(* Logix 5000 project; controller R400_500_XLS vendor 1 type 14 code 216 rev 31.11; software revision 31.01; part 11 of 32 *)
(* tags used below, declared in another part *)
   CalCond : SINT;
   CalFrinseCond : SINT;
   CalibCondCnt : SINT;
   CalibData : UDT_SCALE[8];
   CalibFrinseCondCnt : SINT;
   CalibIndex : DINT;   // Calibration Pointer
   CalibPressCnt : SINT;
   CalPressure : SINT;
   DX_div_100 : REAL;
   M : DINT[5];   // Memory Bits
   ONS_FC86 : DINT;
   rBuffer : REAL[4];
   Supervisor : DINT;
   ChemCond : REAL;
   FinalRinseCond : REAL;
   I_Chem_Cond : DINT;   // Chemical water conductivity
   I_Final_Rinse_Cond : DINT;   // Final rinse water conductivity
   I_Pump_Press : DINT;   // Recirculation pump pressure
   Msg_CalibChem : SINT;
   Msg_CalibFrinse : SINT;
   Msg_CalibPress : SINT;
   Msg_EditCalib : SINT;   // Screen 103 Msg Display
   NumInput : UDT_NUMERIC_INPUT[65];   // Numeric input
   NumInputReal : UDT_NUMERIC_INPUT_REAL[17];
   PmpPres : REAL;
   PressureUnit : BOOL;   // Pressure Unit 0=PSIG 1=BAR
   Screen_Ctrl : DINT;   // PLC Screen Request
   Tpb : DINT[11];
   TpbImage : DINT[11];
   Unit : Hrdwre;   // Unit Configuration
(* MainProgram, continued *)

ROUTINE SPV_10_ANALOG_CHANNEL_CALIBRATION   (* ladder *)
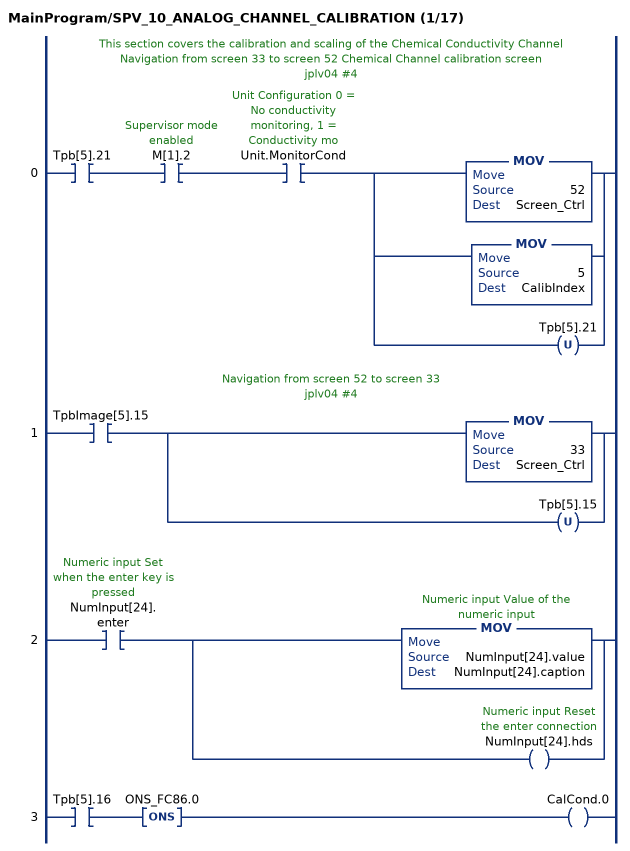
   // This section covers the calibration and scaling of the Chemical Conductivity Channel
   // Navigation from screen 33 to screen 52 Chemical Channel calibration screen
   // jplv04 #4
   0: XIC(Tpb[5].21)XIC(M[1].2)XIC(Unit.MonitorCond)[MOV(52,Screen_Ctrl) ,MOV(5,CalibIndex) ,OTU(Tpb[5].21) ];
   // Navigation from screen 52 to screen 33
   // jplv04 #4
   1: XIC(TpbImage[5].15)[MOV(33,Screen_Ctrl) ,OTU(Tpb[5].15) ];
   2: XIC(NumInput[24].enter)[MOV(NumInput[24].value,NumInput[24].caption) ,OTE(NumInput[24].hds) ];
   3: XIC(Tpb[5].16)ONS(ONS_FC86.0)OTE(CalCond.0);
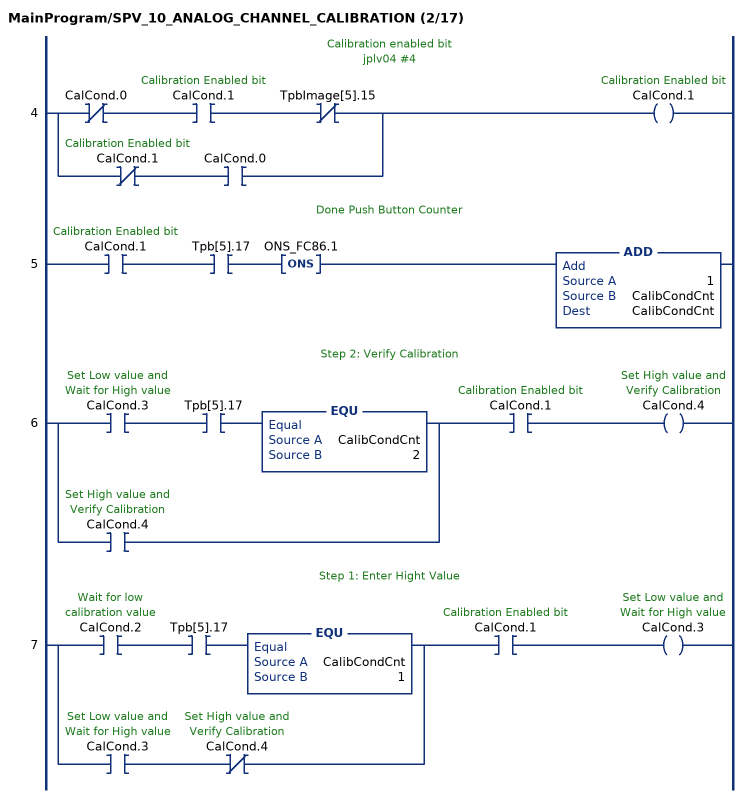
   // Calibration enabled bit
   // jplv04 #4
   4: [XIO(CalCond.0) XIC(CalCond.1) XIO(TpbImage[5].15) ,XIO(CalCond.1) XIC(CalCond.0) ]OTE(CalCond.1);
   // Done Push Button Counter
   5: XIC(CalCond.1)XIC(Tpb[5].17)ONS(ONS_FC86.1)ADD(1,CalibCondCnt,CalibCondCnt);
   // Step 2: Verify Calibration
   6: [XIC(CalCond.3) XIC(Tpb[5].17) EQU(CalibCondCnt,2) ,XIC(CalCond.4) ]XIC(CalCond.1)OTE(CalCond.4);
   // Step 1: Enter Hight Value
   7: [XIC(CalCond.2) XIC(Tpb[5].17) EQU(CalibCondCnt,1) ,XIC(CalCond.3) XIO(CalCond.4) ]XIC(CalCond.1)OTE(CalCond.3);
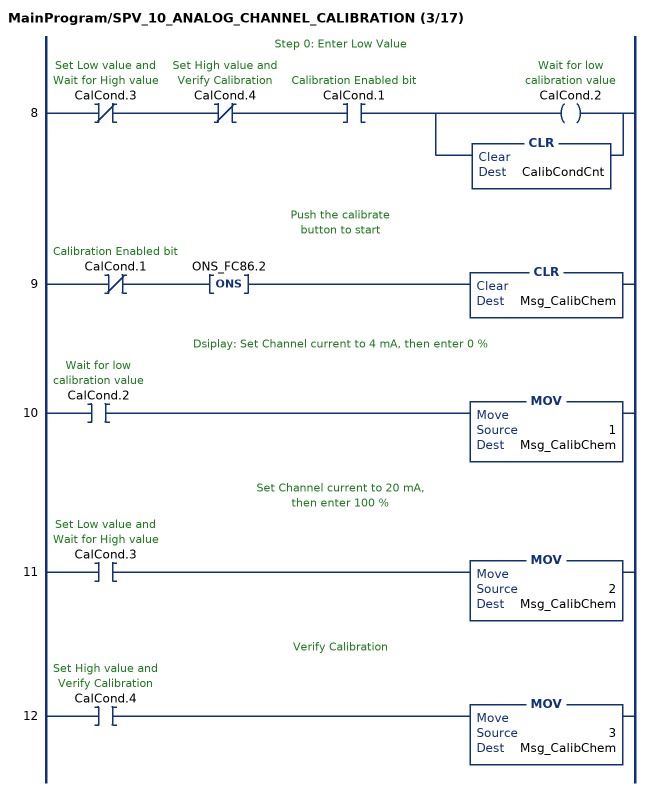
   // Step 0: Enter Low Value
   8: XIO(CalCond.3)XIO(CalCond.4)XIC(CalCond.1)[OTE(CalCond.2) ,CLR(CalibCondCnt) ];
   // Push the calibrate
   // button to start
   9: XIO(CalCond.1)ONS(ONS_FC86.2)CLR(Msg_CalibChem);
   // Dsiplay: Set Channel current to 4 mA, then enter 0 %
   10: XIC(CalCond.2)MOV(1,Msg_CalibChem);
   // Set Channel current to 20 mA,
   // then enter 100 %
   11: XIC(CalCond.3)MOV(2,Msg_CalibChem);
   // Verify Calibration
   12: XIC(CalCond.4)MOV(3,Msg_CalibChem);
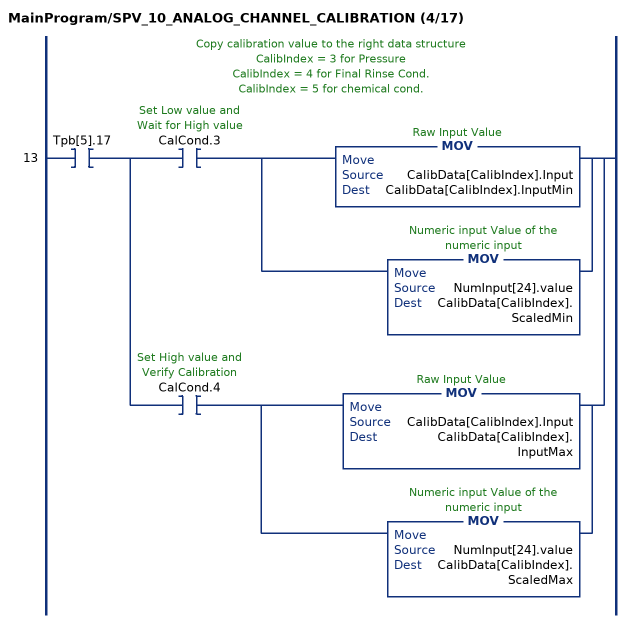
   // Copy calibration value to the right data structure
   // CalibIndex = 3 for Pressure
   // CalibIndex = 4 for Final Rinse Cond.
   // CalibIndex = 5 for chemical cond.
   13: XIC(Tpb[5].17)[XIC(CalCond.3) [MOV(CalibData[CalibIndex].Input,CalibData[CalibIndex].InputMin) ,MOV(NumInput[24].value,CalibData[CalibIndex].ScaledMin) ] ,XIC(CalCond.4) [MOV(CalibData[CalibIndex].Input,CalibData[CalibIndex].InputMax) ,MOV(NumInput[24].value,CalibData[CalibIndex].ScaledMax) ] ];
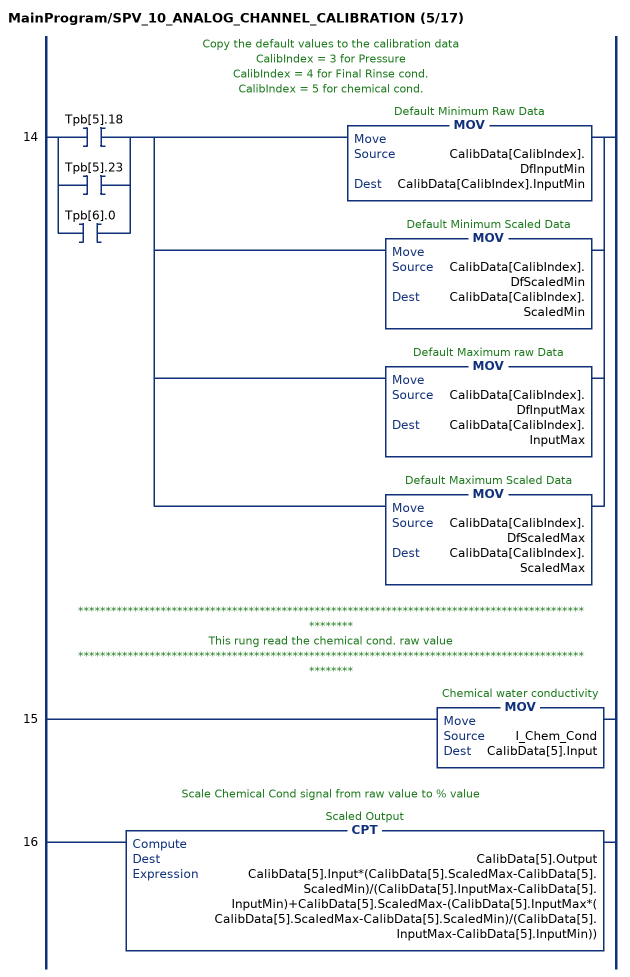
   // Copy the default values to the calibration data
   // CalibIndex = 3 for Pressure
   // CalibIndex = 4 for Final Rinse cond.
   // CalibIndex = 5 for chemical cond.
   14: [XIC(Tpb[5].18) ,XIC(Tpb[5].23) ,XIC(Tpb[6].0) ][MOV(CalibData[CalibIndex].DfInputMin,CalibData[CalibIndex].InputMin) ,MOV(CalibData[CalibIndex].DfScaledMin,CalibData[CalibIndex].ScaledMin) ,MOV(CalibData[CalibIndex].DfInputMax,CalibData[CalibIndex].InputMax) ,MOV(CalibData[CalibIndex].DfScaledMax,CalibData[CalibIndex].ScaledMax) ];
   // ****************************************************************************************************
   // This rung read the chemical cond. raw value
   // ****************************************************************************************************
   15: MOV(I_Chem_Cond,CalibData[5].Input);
   // Scale Chemical Cond signal from raw value to % value
   16: CPT(CalibData[5].Output,CalibData[5].Input*(CalibData[5].ScaledMax-CalibData[5].ScaledMin)/(CalibData[5].InputMax-CalibData[5].InputMin)+CalibData[5].ScaledMax-(CalibData[5].InputMax*(CalibData[5].ScaledMax-CalibData[5].ScaledMin)/(CalibData[5].InputMax-CalibData[5].InputMin)));
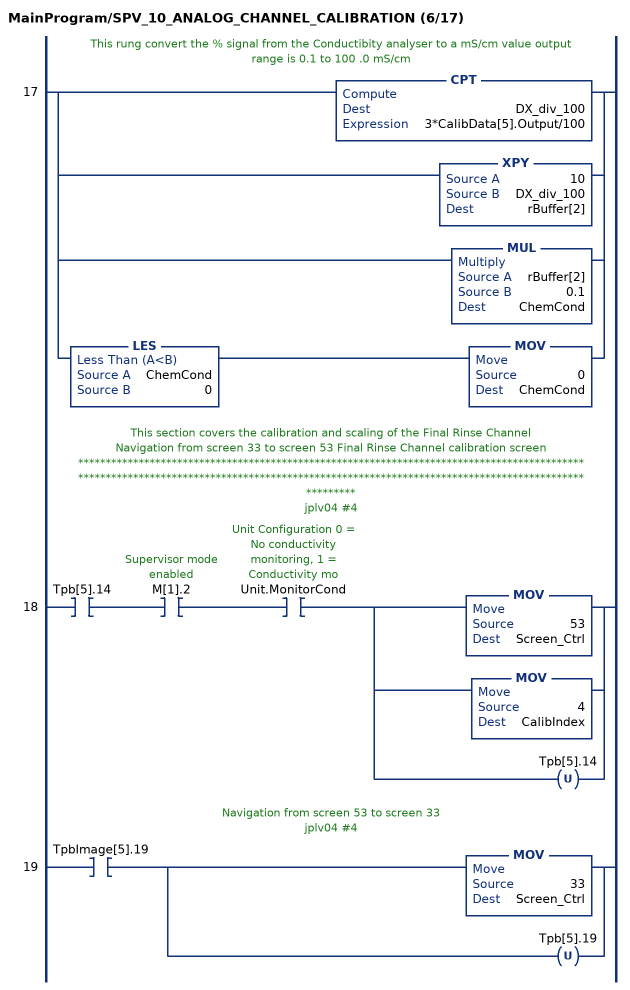
   // This rung convert the % signal from the Conductibity analyser to a mS/cm value output range is 0.1 to 100 .0 mS/cm
   17: [CPT(DX_div_100,3*CalibData[5].Output/100) ,XPY(10,DX_div_100,rBuffer[2]) ,MUL(rBuffer[2],0.1,ChemCond) ,LES(ChemCond,0) MOV(0,ChemCond) ];
   // This section covers the calibration and scaling of the Final Rinse Channel
   // Navigation from screen 33 to screen 53 Final Rinse Channel calibration screen
   // *************************************************************************************************************************************************************************************************
   // jplv04 #4
   18: XIC(Tpb[5].14)XIC(M[1].2)XIC(Unit.MonitorCond)[MOV(53,Screen_Ctrl) ,MOV(4,CalibIndex) ,OTU(Tpb[5].14) ];
   // Navigation from screen 53 to screen 33
   // jplv04 #4
   19: XIC(TpbImage[5].19)[MOV(33,Screen_Ctrl) ,OTU(Tpb[5].19) ];
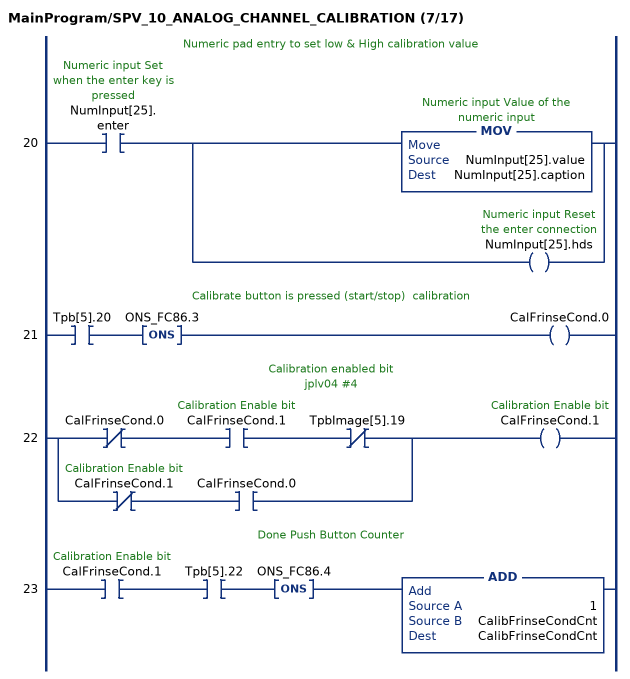
   // Numeric pad entry to set low & High calibration value
   20: XIC(NumInput[25].enter)[MOV(NumInput[25].value,NumInput[25].caption) ,OTE(NumInput[25].hds) ];
   // Calibrate button is pressed (start/stop)  calibration
   21: XIC(Tpb[5].20)ONS(ONS_FC86.3)OTE(CalFrinseCond.0);
   // Calibration enabled bit
   // jplv04 #4
   22: [XIO(CalFrinseCond.0) XIC(CalFrinseCond.1) XIO(TpbImage[5].19) ,XIO(CalFrinseCond.1) XIC(CalFrinseCond.0) ]OTE(CalFrinseCond.1);
   // Done Push Button Counter
   23: XIC(CalFrinseCond.1)XIC(Tpb[5].22)ONS(ONS_FC86.4)ADD(1,CalibFrinseCondCnt,CalibFrinseCondCnt);
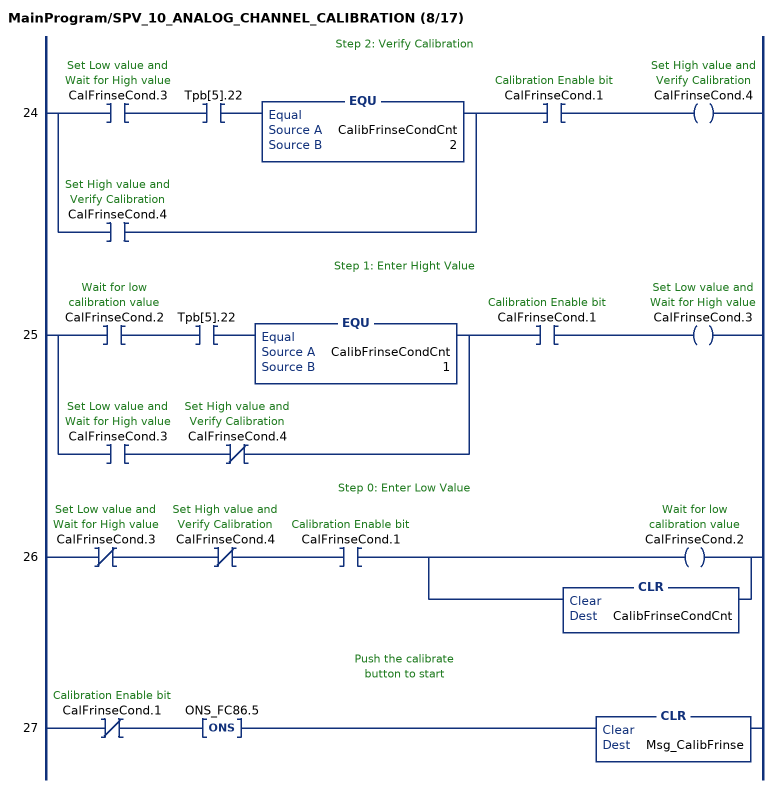
   // Step 2: Verify Calibration
   24: [XIC(CalFrinseCond.3) XIC(Tpb[5].22) EQU(CalibFrinseCondCnt,2) ,XIC(CalFrinseCond.4) ]XIC(CalFrinseCond.1)OTE(CalFrinseCond.4);
   // Step 1: Enter Hight Value
   25: [XIC(CalFrinseCond.2) XIC(Tpb[5].22) EQU(CalibFrinseCondCnt,1) ,XIC(CalFrinseCond.3) XIO(CalFrinseCond.4) ]XIC(CalFrinseCond.1)OTE(CalFrinseCond.3);
   // Step 0: Enter Low Value
   26: XIO(CalFrinseCond.3)XIO(CalFrinseCond.4)XIC(CalFrinseCond.1)[OTE(CalFrinseCond.2) ,CLR(CalibFrinseCondCnt) ];
   // Push the calibrate
   // button to start
   27: XIO(CalFrinseCond.1)ONS(ONS_FC86.5)CLR(Msg_CalibFrinse);
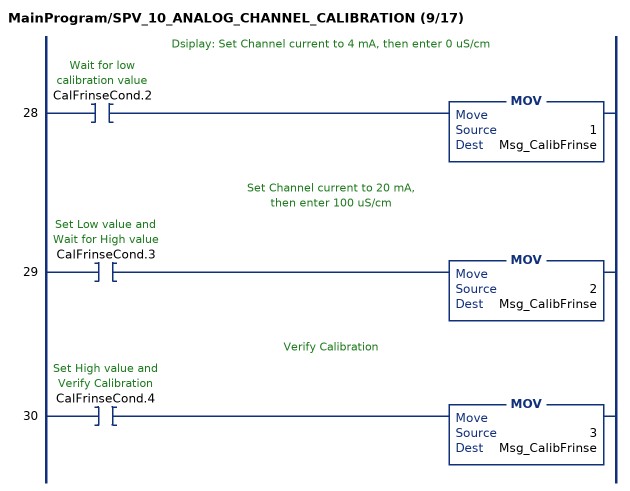
   // Dsiplay: Set Channel current to 4 mA, then enter 0 uS/cm
   28: XIC(CalFrinseCond.2)MOV(1,Msg_CalibFrinse);
   // Set Channel current to 20 mA,
   // then enter 100 uS/cm
   29: XIC(CalFrinseCond.3)MOV(2,Msg_CalibFrinse);
   // Verify Calibration
   30: XIC(CalFrinseCond.4)MOV(3,Msg_CalibFrinse);
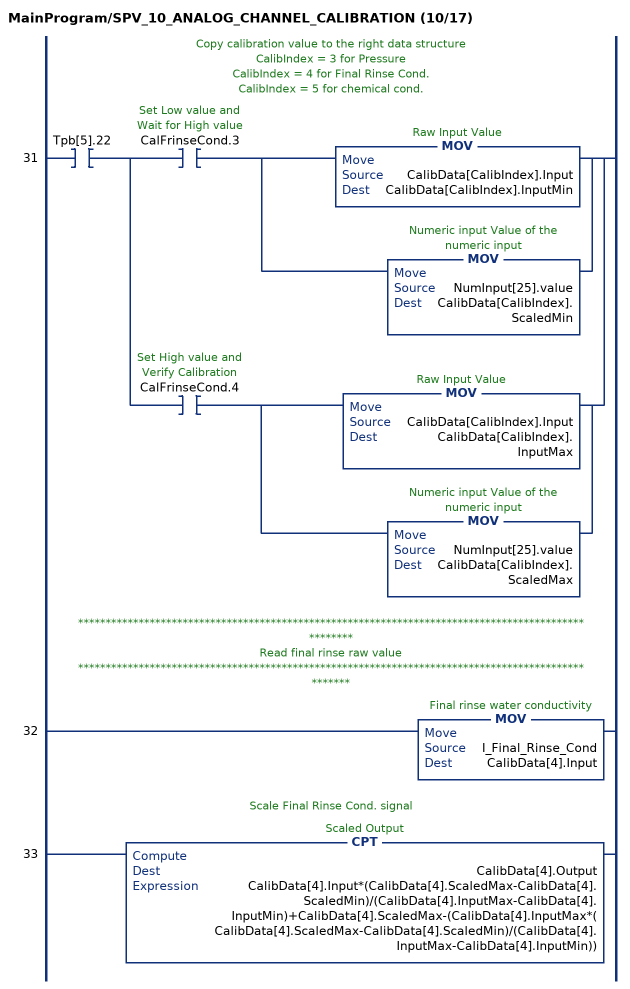
   // Copy calibration value to the right data structure
   // CalibIndex = 3 for Pressure
   // CalibIndex = 4 for Final Rinse Cond.
   // CalibIndex = 5 for chemical cond.
   31: XIC(Tpb[5].22)[XIC(CalFrinseCond.3) [MOV(CalibData[CalibIndex].Input,CalibData[CalibIndex].InputMin) ,MOV(NumInput[25].value,CalibData[CalibIndex].ScaledMin) ] ,XIC(CalFrinseCond.4) [MOV(CalibData[CalibIndex].Input,CalibData[CalibIndex].InputMax) ,MOV(NumInput[25].value,CalibData[CalibIndex].ScaledMax) ] ];
   // ****************************************************************************************************
   // Read final rinse raw value
   // ***************************************************************************************************
   32: MOV(I_Final_Rinse_Cond,CalibData[4].Input);
   // Scale Final Rinse Cond. signal
   33: CPT(CalibData[4].Output,CalibData[4].Input*(CalibData[4].ScaledMax-CalibData[4].ScaledMin)/(CalibData[4].InputMax-CalibData[4].InputMin)+CalibData[4].ScaledMax-(CalibData[4].InputMax*(CalibData[4].ScaledMax-CalibData[4].ScaledMin)/(CalibData[4].InputMax-CalibData[4].InputMin)));
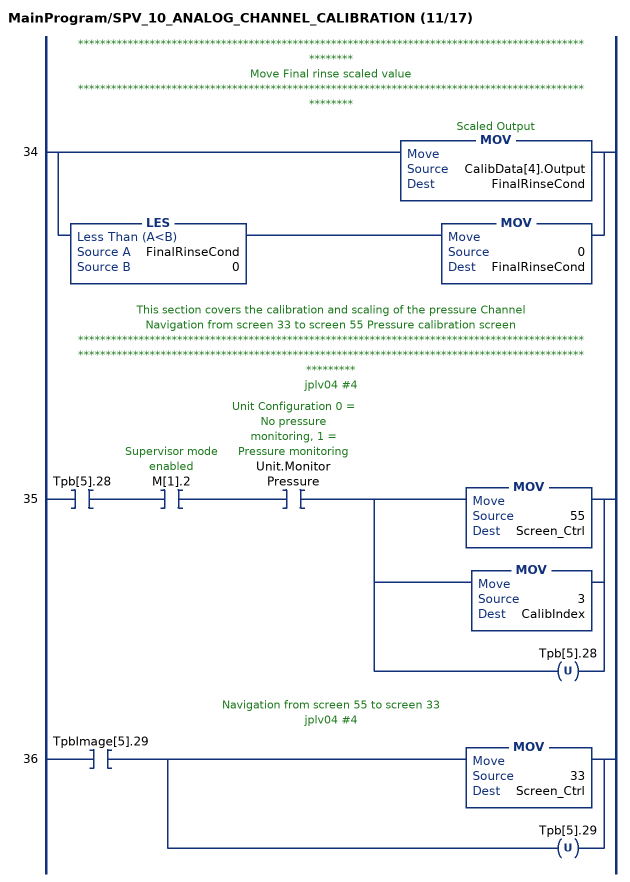
   // ****************************************************************************************************
   // Move Final rinse scaled value
   // ****************************************************************************************************
   34: [MOV(CalibData[4].Output,FinalRinseCond) ,LES(FinalRinseCond,0) MOV(0,FinalRinseCond) ];
   // This section covers the calibration and scaling of the pressure Channel
   // Navigation from screen 33 to screen 55 Pressure calibration screen
   // *************************************************************************************************************************************************************************************************
   // jplv04 #4
   35: XIC(Tpb[5].28)XIC(M[1].2)XIC(Unit.MonitorPressure)[MOV(55,Screen_Ctrl) ,MOV(3,CalibIndex) ,OTU(Tpb[5].28) ];
   // Navigation from screen 55 to screen 33
   // jplv04 #4
   36: XIC(TpbImage[5].29)[MOV(33,Screen_Ctrl) ,OTU(Tpb[5].29) ];
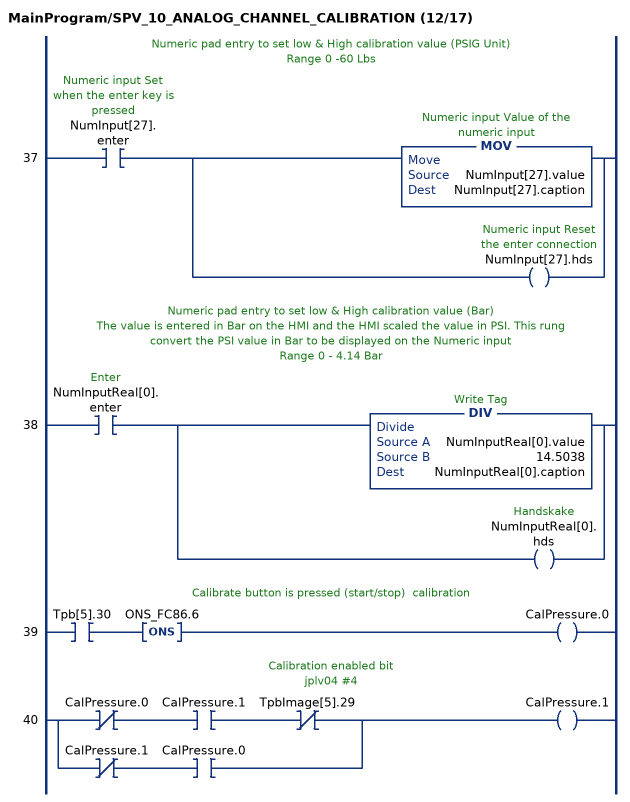
   // Numeric pad entry to set low & High calibration value (PSIG Unit)
   // Range 0 -60 Lbs
   37: XIC(NumInput[27].enter)[MOV(NumInput[27].value,NumInput[27].caption) ,OTE(NumInput[27].hds) ];
   // Numeric pad entry to set low & High calibration value (Bar)
   // The value is entered in Bar on the HMI and the HMI scaled the value in PSI. This rung convert the PSI value in Bar to be displayed on the Numeric input
   // Range 0 - 4.14 Bar
   38: XIC(NumInputReal[0].enter)[DIV(NumInputReal[0].value,14.5038,NumInputReal[0].caption) ,OTE(NumInputReal[0].hds) ];
   // Calibrate button is pressed (start/stop)  calibration
   39: XIC(Tpb[5].30)ONS(ONS_FC86.6)OTE(CalPressure.0);
   // Calibration enabled bit
   // jplv04 #4
   40: [XIO(CalPressure.0) XIC(CalPressure.1) XIO(TpbImage[5].29) ,XIO(CalPressure.1) XIC(CalPressure.0) ]OTE(CalPressure.1);
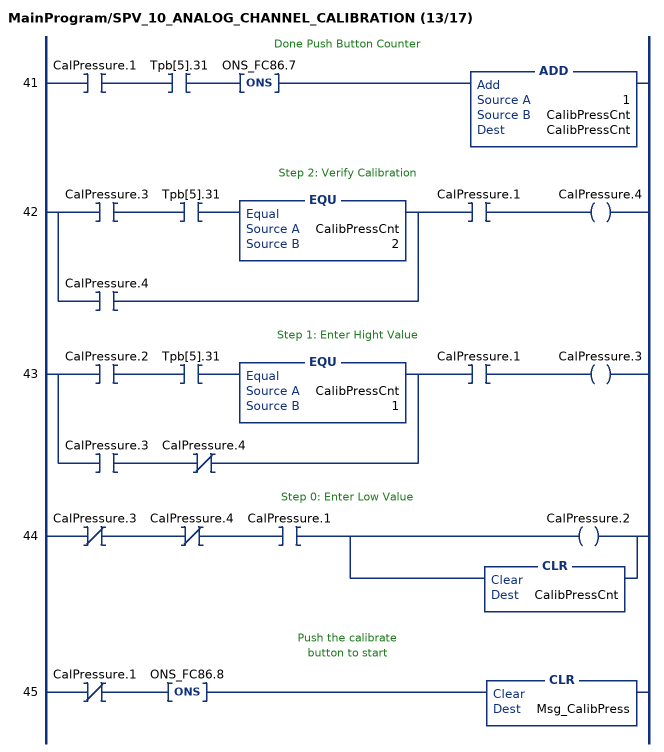
   // Done Push Button Counter
   41: XIC(CalPressure.1)XIC(Tpb[5].31)ONS(ONS_FC86.7)ADD(1,CalibPressCnt,CalibPressCnt);
   // Step 2: Verify Calibration
   42: [XIC(CalPressure.3) XIC(Tpb[5].31) EQU(CalibPressCnt,2) ,XIC(CalPressure.4) ]XIC(CalPressure.1)OTE(CalPressure.4);
   // Step 1: Enter Hight Value
   43: [XIC(CalPressure.2) XIC(Tpb[5].31) EQU(CalibPressCnt,1) ,XIC(CalPressure.3) XIO(CalPressure.4) ]XIC(CalPressure.1)OTE(CalPressure.3);
   // Step 0: Enter Low Value
   44: XIO(CalPressure.3)XIO(CalPressure.4)XIC(CalPressure.1)[OTE(CalPressure.2) ,CLR(CalibPressCnt) ];
   // Push the calibrate
   // button to start
   45: XIO(CalPressure.1)ONS(ONS_FC86.8)CLR(Msg_CalibPress);
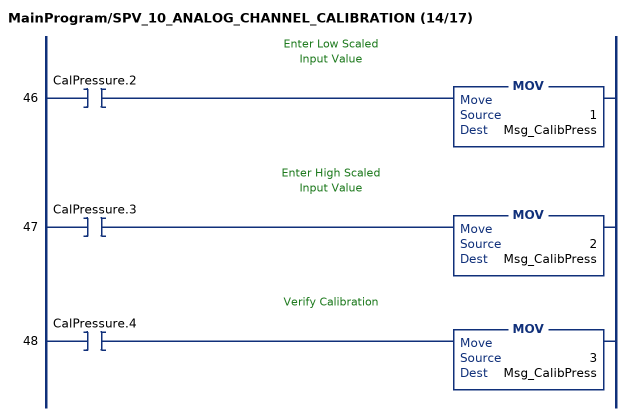
   // Enter Low Scaled
   // Input Value
   46: XIC(CalPressure.2)MOV(1,Msg_CalibPress);
   // Enter High Scaled
   // Input Value
   47: XIC(CalPressure.3)MOV(2,Msg_CalibPress);
   // Verify Calibration
   48: XIC(CalPressure.4)MOV(3,Msg_CalibPress);
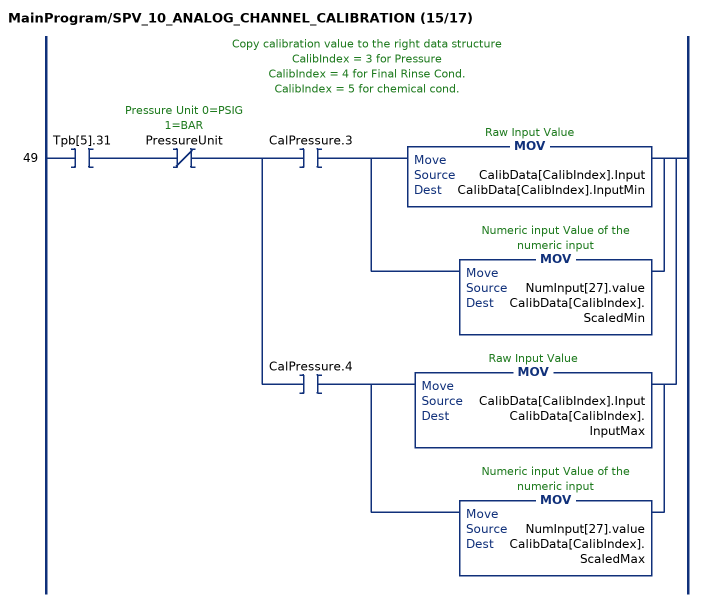
   // Copy calibration value to the right data structure
   // CalibIndex = 3 for Pressure
   // CalibIndex = 4 for Final Rinse Cond.
   // CalibIndex = 5 for chemical cond.
   49: XIC(Tpb[5].31)XIO(PressureUnit)[XIC(CalPressure.3) [MOV(CalibData[CalibIndex].Input,CalibData[CalibIndex].InputMin) ,MOV(NumInput[27].value,CalibData[CalibIndex].ScaledMin) ] ,XIC(CalPressure.4) [MOV(CalibData[CalibIndex].Input,CalibData[CalibIndex].InputMax) ,MOV(NumInput[27].value,CalibData[CalibIndex].ScaledMax) ] ];
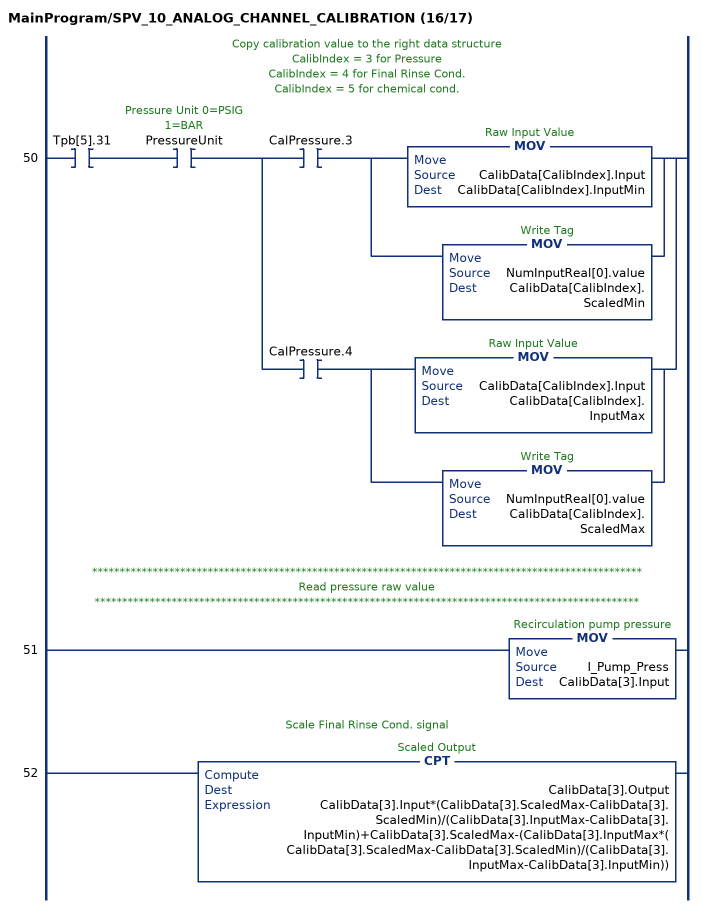
   // Copy calibration value to the right data structure
   // CalibIndex = 3 for Pressure
   // CalibIndex = 4 for Final Rinse Cond.
   // CalibIndex = 5 for chemical cond.
   50: XIC(Tpb[5].31)XIC(PressureUnit)[XIC(CalPressure.3) [MOV(CalibData[CalibIndex].Input,CalibData[CalibIndex].InputMin) ,MOV(NumInputReal[0].value,CalibData[CalibIndex].ScaledMin) ] ,XIC(CalPressure.4) [MOV(CalibData[CalibIndex].Input,CalibData[CalibIndex].InputMax) ,MOV(NumInputReal[0].value,CalibData[CalibIndex].ScaledMax) ] ];
   // ****************************************************************************************************
   // Read pressure raw value
   // ***************************************************************************************************
   51: MOV(I_Pump_Press,CalibData[3].Input);
   // Scale Final Rinse Cond. signal
   52: CPT(CalibData[3].Output,CalibData[3].Input*(CalibData[3].ScaledMax-CalibData[3].ScaledMin)/(CalibData[3].InputMax-CalibData[3].InputMin)+CalibData[3].ScaledMax-(CalibData[3].InputMax*(CalibData[3].ScaledMax-CalibData[3].ScaledMin)/(CalibData[3].InputMax-CalibData[3].InputMin)));
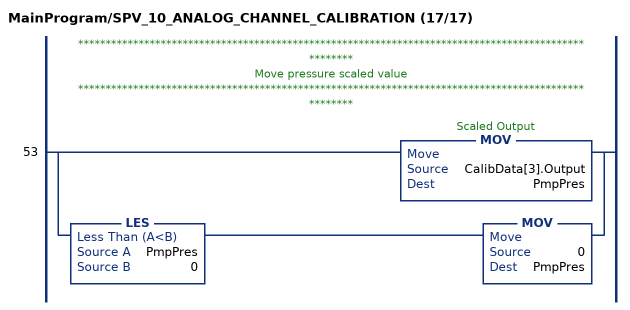
   // ****************************************************************************************************
   // Move pressure scaled value
   // ****************************************************************************************************
   53: [MOV(CalibData[3].Output,PmpPres) ,LES(PmpPres,0) MOV(0,PmpPres) ];
END_ROUTINE

ROUTINE SPV_11_EDIT_CALIBRATION   (* ladder *)
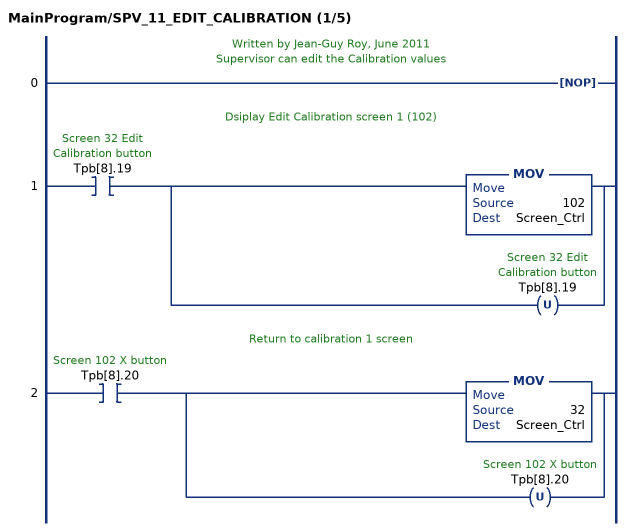
   // Written by Jean-Guy Roy, June 2011
   // Supervisor can edit the Calibration values
   0: NOP();
   // Dsiplay Edit Calibration screen 1 (102)
   1: XIC(Tpb[8].19)[MOV(102,Screen_Ctrl) ,OTU(Tpb[8].19) ];
   // Return to calibration 1 screen
   2: XIC(Tpb[8].20)[MOV(32,Screen_Ctrl) ,OTU(Tpb[8].20) ];
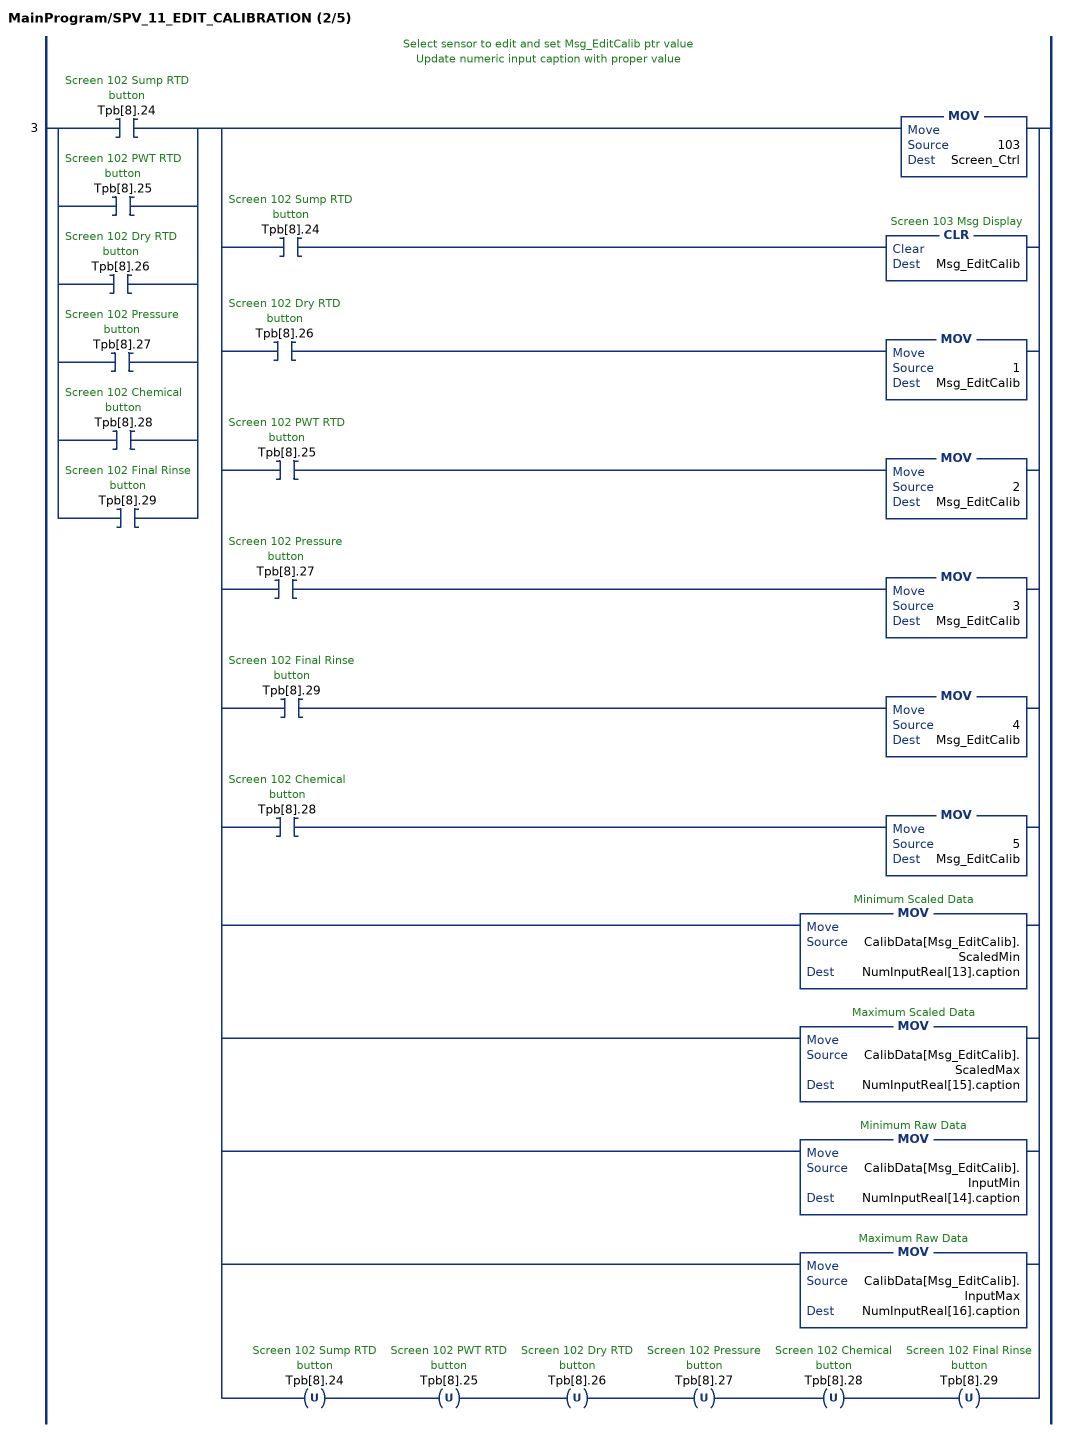
   // Select sensor to edit and set Msg_EditCalib ptr value
   // Update numeric input caption with proper value
   3: [XIC(Tpb[8].24) ,XIC(Tpb[8].25) ,XIC(Tpb[8].26) ,XIC(Tpb[8].27) ,XIC(Tpb[8].28) ,XIC(Tpb[8].29) ][MOV(103,Screen_Ctrl) ,XIC(Tpb[8].24) CLR(Msg_EditCalib) ,XIC(Tpb[8].26) MOV(1,Msg_EditCalib) ,XIC(Tpb[8].25) MOV(2,Msg_EditCalib) ,XIC(Tpb[8].27) MOV(3,Msg_EditCalib) ,XIC(Tpb[8].29) MOV(4,Msg_EditCalib) ,XIC(Tpb[8].28) MOV(5,Msg_EditCalib) ,MOV(CalibData[Msg_EditCalib].ScaledMin,NumInputReal[13].caption) ,MOV(CalibData[Msg_EditCalib].ScaledMax,NumInputReal[15].caption) ,MOV(CalibData[Msg_EditCalib].InputMin,NumInputReal[14].caption) ,MOV(CalibData[Msg_EditCalib].InputMax,NumInputReal[16].caption) ,OTU(Tpb[8].24) OTU(Tpb[8].25) OTU(Tpb[8].26) OTU(Tpb[8].27) OTU(Tpb[8].28) OTU(Tpb[8].29) ];
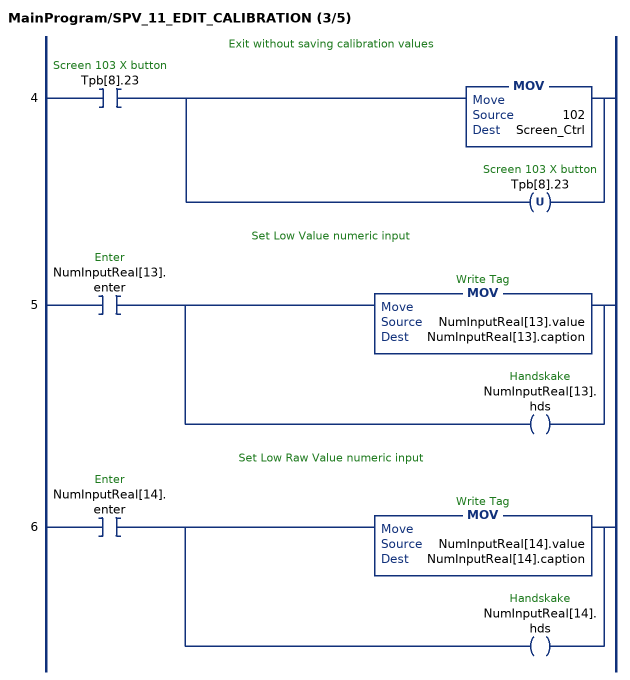
   // Exit without saving calibration values
   4: XIC(Tpb[8].23)[MOV(102,Screen_Ctrl) ,OTU(Tpb[8].23) ];
   // Set Low Value numeric input
   5: XIC(NumInputReal[13].enter)[MOV(NumInputReal[13].value,NumInputReal[13].caption) ,OTE(NumInputReal[13].hds) ];
   // Set Low Raw Value numeric input
   6: XIC(NumInputReal[14].enter)[MOV(NumInputReal[14].value,NumInputReal[14].caption) ,OTE(NumInputReal[14].hds) ];
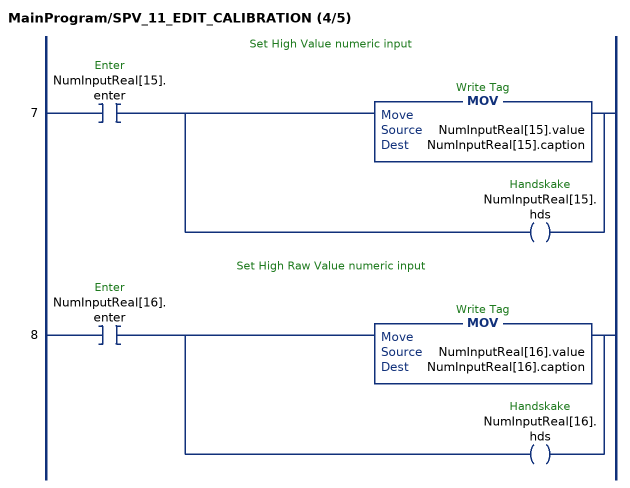
   // Set High Value numeric input
   7: XIC(NumInputReal[15].enter)[MOV(NumInputReal[15].value,NumInputReal[15].caption) ,OTE(NumInputReal[15].hds) ];
   // Set High Raw Value numeric input
   8: XIC(NumInputReal[16].enter)[MOV(NumInputReal[16].value,NumInputReal[16].caption) ,OTE(NumInputReal[16].hds) ];
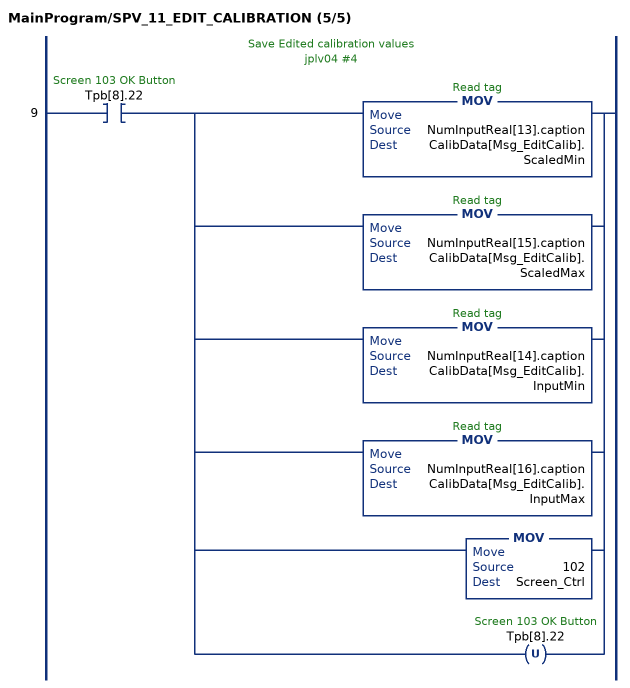
   // Save Edited calibration values
   // jplv04 #4
   9: XIC(Tpb[8].22)[MOV(NumInputReal[13].caption,CalibData[Msg_EditCalib].ScaledMin) ,MOV(NumInputReal[15].caption,CalibData[Msg_EditCalib].ScaledMax) ,MOV(NumInputReal[14].caption,CalibData[Msg_EditCalib].InputMin) ,MOV(NumInputReal[16].caption,CalibData[Msg_EditCalib].InputMax) ,MOV(102,Screen_Ctrl) ,OTU(Tpb[8].22) ];
END_ROUTINE
